VAR_GLOBAL
    // PLC 内部手动命令与轴反馈；命令由 A03_ManualCommands 转交，反馈由基础轴块更新。
    // 上位机手动命令写 GVL_control.aStation[站号].aAxis，状态读取 GVL_HMI.stMonitor。

    Axis1 : ST_AxisAds; // 轴1内部手动命令与实际反馈；命令由命令门转交，反馈由轴1基础块更新。
    Axis2 : ST_AxisAds; // 轴2内部手动命令与实际反馈；命令由命令门转交，反馈由轴2基础块更新。
    Axis3 : ST_AxisAds; // 轴3内部手动命令与实际反馈；命令由命令门转交，反馈由轴3基础块更新。
    Axis4 : ST_AxisAds; // 轴4内部手动命令与实际反馈；命令由命令门转交，反馈由轴4基础块更新。


END_VAR

(* stored: Version 1.1.0.1
   GVL GVL_axis: Id {26300288-3096-43e2-833c-dddff8221f5e} *)
